(* IEC 61131-3 sources: plc-iiot-stack/src/POUs/Iiot/F_IiotAlarmStateText, 2 files *)

(* ---- F_IiotAlarmStateText.decl.st ---- *)
// Назначение: имя состояния тревоги для полей state и prev_state.
// Автор:      kr0nsch
// Версия:     0.1.0
// Документ:   docs/plc_mqtt.md, раздел «Тревоги»
FUNCTION F_IiotAlarmStateText : STRING(GVL_Const.IIOT_TEXT_LEN)
VAR_INPUT
    eState : E_IiotAlarmState;
END_VAR

(* ---- F_IiotAlarmStateText.impl.st ---- *)
CASE eState OF
    E_IiotAlarmState.Normal:
        F_IiotAlarmStateText := 'Normal';
    E_IiotAlarmState.ActiveUnack:
        F_IiotAlarmStateText := 'ActiveUnack';
    E_IiotAlarmState.ActiveAck:
        F_IiotAlarmStateText := 'ActiveAck';
    E_IiotAlarmState.RtnUnack:
        F_IiotAlarmStateText := 'RtnUnack';
    E_IiotAlarmState.Shelved:
        F_IiotAlarmStateText := 'Shelved';
    E_IiotAlarmState.SuppressedByDesign:
        F_IiotAlarmStateText := 'SuppressedByDesign';
ELSE
    F_IiotAlarmStateText := 'OutOfService';
END_CASE
